{attribute 'linkalways'} 
{attribute 'no_explicit_call' := 'This FB is a CLASS and must be accessed using methods or properties'}
{attribute 'enable_dynamic_creation'}
FUNCTION_BLOCK _ETcVnCalibrationPattern EXTENDS EnumDatatypeBase
VAR
	localData : ETcVnCalibrationPattern;
	activeData : REFERENCE TO ETcVnCalibrationPattern;
	enumBaseDatatype : _DINT(localData);
END_VAR

METHOD PRIVATE AddLocalEnumeration
VAR_INPUT
	Enumeration : T_MAXSTRING;
	Value : ETcVnCalibrationPattern;
END_VAR
AddEnumeration(Enumeration, Value);
END_METHOD

PROPERTY PUBLIC Address : PVOID
GET
Address := ADR(activeData);
END_GET
END_PROPERTY

METHOD PUBLIC ClearReference
VAR_INPUT
END_VAR
activeData REF= localData;
SetBaseDatatypeReference();
END_METHOD

METHOD PUBLIC Clone : I_Datatype
VAR
    pClone : POINTER TO _ETcVnCalibrationPattern;
END_VAR
pClone := __NEW(_ETcVnCalibrationPattern(InitialValue := Value));
Clone := pClone^;
END_METHOD

METHOD FB_init : BOOL
VAR_INPUT
	bInitRetains : BOOL; // if TRUE, the retain variables are initialized (warm start / cold start)
	bInCopyCode : BOOL;  // if TRUE, the instance afterwards gets moved into the copy code (online change)
	InitialValue : ETcVnCalibrationPattern;
END_VAR
localData := InitialValue;
AddBaseDatatype(enumBaseDatatype);
ClearReference();

AddLocalEnumeration('TCVN_CP_CIRCLES_SYM', ETcVnCalibrationPattern.TCVN_CP_CIRCLES_SYM);
AddLocalEnumeration('TCVN_CP_CIRCLES_ASYM', ETcVnCalibrationPattern.TCVN_CP_CIRCLES_ASYM);
AddLocalEnumeration('TCVN_CP_CIRCLES_ASYM_INDENT', ETcVnCalibrationPattern.TCVN_CP_CIRCLES_ASYM_INDENT);
END_METHOD

PROPERTY PUBLIC Identifier : T_MAXSTRING
GET
Identifier := 'ETcVnCalibrationPattern';
END_GET
END_PROPERTY

METHOD IsEnumeratorValueEqual : BOOL
VAR_INPUT
	Enumerator : I_KeyValueForwardEnumerator;
END_VAR
VAR
	storedValue : ETcVnCalibrationPattern;
END_VAR
IF NOT Enumerator.TryGet(storedValue) THEN
	RETURN;
END_IF

IsEnumeratorValueEqual := storedValue = activeData;
END_METHOD

METHOD PUBLIC MakeReferenceTo
VAR_INPUT
	ReferenceTarget : REFERENCE TO ETcVnCalibrationPattern;
END_VAR
activeData REF= ReferenceTarget;
SetBaseDatatypeReference();
END_METHOD

METHOD PROTECTED SetBaseDatatypeReference
VAR_INPUT
END_VAR
enumBaseDatatype.MakeReferenceTo(activeData);
END_METHOD

PROPERTY PUBLIC Size : UDINT
GET
Size := SIZEOF(activeData);
END_GET
END_PROPERTY

METHOD TryMakeReferenceTo : BOOL
VAR_INPUT
	Target : I_Datatype;
END_VAR
VAR
	pTargetData : POINTER TO ETcVnCalibrationPattern;
END_VAR
IF NOT IsEquivalentTo(Target) THEN
	RETURN;
END_IF

pTargetData := Target.Address;
activeData REF= pTargetData^;
SetBaseDatatypeReference();
TryMakeReferenceTo := TRUE;
END_METHOD

PROPERTY PUBLIC Value : ETcVnCalibrationPattern
GET
Value := activeData;
END_GET
SET
activeData := Value;
END_SET
END_PROPERTY

END_FUNCTION_BLOCK

(* stored: Version 1.1.0.1, ProductVersion 3.1.4024.13
   POU _ETcVnCalibrationPattern: Id {242b7478-690d-4c28-ab58-0771f86f04d1}, SpecialFunc None
   Folder Core: Id {89ac6c03-fe2b-0412-3140-ce12b5294cca}
   Folder Protected: Id {3e24fde9-72a3-066e-33f7-db344d163029}
   Folder Customize: Id {7ec4a401-f658-022c-09dd-eb1a8780c610}
   Folder Constructor: Id {052bf58e-5e75-4250-8666-3b9d80163253}
   Folder Private: Id {96d89ac4-5ec6-4c6f-b6d5-705b3acea75e}
   Folder Protected: Id {c95cf233-58df-454c-b43f-f514fde668b9}
   Method AddLocalEnumeration: Id {27784235-ed37-44c2-ad52-aef4feaedbb7}
   Property Address: Id {f938c40c-458d-0ebe-2d70-ae5a35cd9e6c}
   Get Get: Id {d2a514e3-f53a-05db-3ada-1a206d9e99a3}
   Method ClearReference: Id {9c416157-ff32-00e9-2725-315f76baca62}
   Method Clone: Id {b06a644d-f512-402b-9c78-fa94ca876d2a}
   Method FB_init: Id {41dea6d3-5ac5-4887-8e07-4c2e9d3d334f}
   Property Identifier: Id {cf6ce56b-f9fb-4e8f-bcf4-45eb1baf4ca7}
   Get Get: Id {d637b286-1d02-4673-8d31-208312ec9c14}
   Method IsEnumeratorValueEqual: Id {36c49053-c56a-4947-8417-32197656628f}
   Method MakeReferenceTo: Id {f5071b5c-f603-42b4-a27f-6f4ff65c1844}
   Method SetBaseDatatypeReference: Id {a669159e-edba-0915-34f5-38d97891b2ca}
   Property Size: Id {0312bbb3-b593-041d-2545-f32b5259207f}
   Get Get: Id {a2c58123-fdad-058f-0376-826f4c97e492}
   Method TryMakeReferenceTo: Id {8ffa0e03-761f-4b19-ad58-7d91491f4e7a}
   Property Value: Id {92425e6b-21c4-400a-892f-54440ae8e267}
   Get Get: Id {bde5f00d-11c9-4d97-894e-2e46c53f46aa}
   Set Set: Id {f7a59fbb-830e-419d-b216-30ba25e1009f} *)
